// TIA Portal V19 export
TYPE "ST_TPM_AutoRecipe"
   STRUCT
      Valid : Bool;
      RecipeId : Int;
      R1Pick { S7_SetPoint := 'True'} : Array[1..4] of "ST_TPM_AutoPosition";
      R1Place { S7_SetPoint := 'True'} : "ST_TPM_AutoPosition";
      R2Pick { S7_SetPoint := 'True'} : "ST_TPM_AutoPosition";
      R2Place { S7_SetPoint := 'True'} : "ST_TPM_AutoPosition";
      R3Pick { S7_SetPoint := 'True'} : "ST_TPM_AutoPosition";
      R3Place { S7_SetPoint := 'True'} : "ST_TPM_AutoPosition";
      StepDistance : LReal;   // Axis engineering units, positive forward.
      StepVelocity : LReal;
      ExitSpeed : Real;   // Engineering units agreed with the drive adapter.
      BeltCapacity : Int;   // Maximum validated number of products on the indexing belt.
      MaxIndexSteps : Int;   // Maximum steps for one product to reach the end.
   END_STRUCT;
END_TYPE
